Staubli VAL3: Force6Item.pjx

--- Force6Item.pjx ---
Parameters version=s8.15.3Cs9_BS3337 stackSize=5000 millimeterUnit=true
Program file=start.pgx
Program file=stop.pgx
Data file=Force6Item.dtx

--- Force6Item.dtx ---
mdesc mNomSpeed
public string sArmType
public num nMaxJnt6Force[6]

--- start.pgx ---
program start()
begin
end

--- stop.pgx ---
program stop()
begin
end
